Universal Robots PolyScope program: AdientTorsF_Eol21.urp

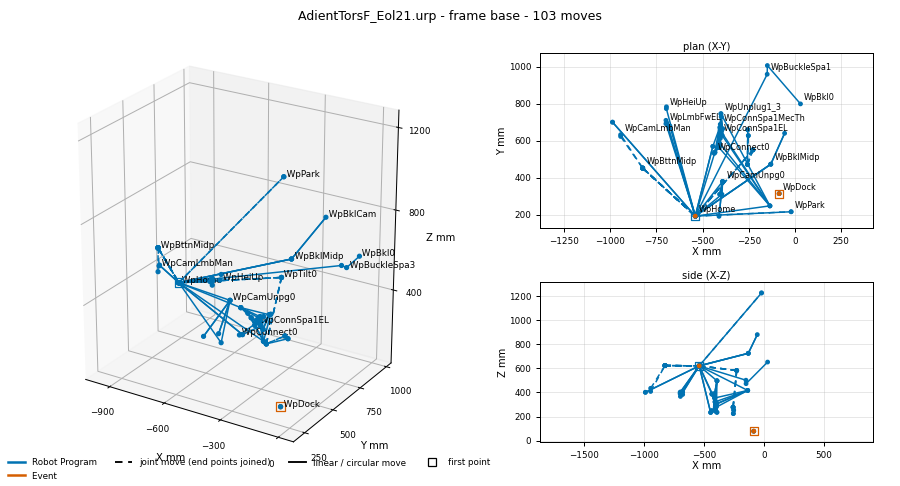
[picture p0: tool path of AdientTorsF_Eol21.urp in frame base, 103 of 155 moves have a stored position in this frame; points joined in program order, loops and branches not executed]
Program AdientTorsF_Eol21 (installation=EOL_21 directory=/programs createdIn=3.5.1 lastSavedIn=5.26.0 robotSerialNumber=20265101890)
Calibrated DH parameters: a=[0.000035, -0.496948, -0.566193, -0.00002, -0.00001, 0]; d=[0.180707, 184.637728, -195.556152, 11.09222, 0.119882, 0.115586]; alpha=[1.570552, -0.001939, 0.006964, 1.570414, -1.570475, 0]; deltaTheta=[0, -0.624231, 6.773924, 0.133492, -0.000002, 0]
InitVariablesNode variables(variable(name=Abort, expression=False), variable(name=AdapterReady, expression=False), variable(name=CMD_Heartbt_i1, expression=0), variable(name=CMD_Program_i1, expression=0), variable(name=CMD_Reserve_i1, expression=0), variable(name=CMD_Timeout_i1, expression=0), variable(name=CamCorrectnOK, expression=0), variable(name=DEBUG, expression=False), variable(name=D_rel, expression=p[0,0,0,0,0,0]), variable(name=EvtBeep, expression=False), variable(name=EvtDock, expression=0), variable(name=Mute, expression=False), variable(name=P_ini, expression=get_actual_tcp_pose()), variable(name=Parking, expression=0), variable(name=ProgExe, expression=0), variable(name=PusherPosFt, expression=0), variable(name=PusherReturn, expression=True), variable(name=STS_Heartbeat, expression=False), variable(name=STS_Progress, expression=0), variable(name=STS_Reservation, expression=0), variable(name=SetCameraProg, expression=0), variable(name=T_KeepReservtn, expression=0), variable(name=Tilt_PV, expression=0))
BeforeStart
  SuppressedNode
    DEBUG := True
  'SW version, to be used to track changes and keep sync of all stations'
  SW_Ver := 1.0
  Folder Scripts [hidden by the author, left out]
  Folder Avoid guidance screen
    Wp := get_actual_tcp_pose()
    MoveJ speed 120 deg/s, acceleration 500 deg/s^2 (useActiveTCP=true optimoveEnabled=false optiMoveSpeed=0.3 optiMoveAcceleration=0.09) feature=Base
      Waypoint Variable (Variable): variable=Wp
  Call GripperOpen
  GoToHome := True
  Script: socket_open("127.0.0.1",30001)
Robot Program (runOnlyOnce=false)
  Folder Execute Program
    Folder Init
      Wait Condition expression=EvtDock≤0
      Folder Verify Adapter ready
        If Di_Docked or AI_Gripper<(ivGripSensOpen+0.3)
          AdapterReady := False
      Folder Go to home pos automatically
        If GoToHome and  not AdapterReady
          Wait Sleep waitTime=1
          If InRange(P_Flange[0],-1,-0.2) and InRange(P_Flange[1],-0.5,0.5) and InRange(P_Flange[2],0.3,1)
            If AdapterDocked or DEBUG or (AI_Gripper<(ivGripSensOpen+0.3))
              MoveJ speed 120 deg/s, acceleration 500 deg/s^2 (useActiveTCP=false positionType=JointAngles optimoveEnabled=false optiMoveSpeed=0.3 optiMoveAcceleration=0.09) tcp=t0_Flange; feature=Base
                Waypoint WpHome: TCP in base x=-539.74 y=192.879 z=621.496 mm, rx=3.1416 ry=0 rz=0 rad; joints [177.915, -76.399, -107.627, -86.021, 90.391, 88.106] deg
            Else 
              Popup Error (haltProgram=false message=Adapter must be docked inputType=Text)
              Halt
          ElseIf AtParkPos
            MoveJ speed 120 deg/s, acceleration 500 deg/s^2 (useActiveTCP=false positionType=JointAngles optimoveEnabled=false optiMoveSpeed=0.3 optiMoveAcceleration=0.09) tcp=t0_Flange; feature=Base
              Waypoint WpPark: TCP in base x=-21.021 y=216.43 z=1228.484 mm, rx=-2.2794 ry=-2.1557 rz=0.0038 rad; joints [148.842, -80.043, -21.696, -168.004, 90.169, -28.26] deg
          Else 
            Popup Error (haltProgram=false message=Illegal position. Adjust arm to open space in front of the backrest, or [Move]->[Home] inputType=Text)
            Halt
        GoToHome := False
      If DEBUG
        'Popup window with program selection'
        ProgExe :=  (valueSource=Operator message=Program number? valueType=Integer)
      If ProgExe>0
        Folder Init
          Mute := False
          Wait Condition expression=not GoToHome
          If not In(ProgExe,[11,12,13,14])
            AdapterReady := False
    Folder Programs
      If InRange(ProgExe,1,99)
        Folder Undock
          If In(ProgExe,[11])
            Script: Report(1)
            If not AdapterReady
              Folder AtHome? [hidden by the author, left out]
              If Progress_run() and  not AdapterDocked
                Script: Report(94)
              If Progress_run()
                Folder Undock
                  MoveL speed 1000 mm/s, acceleration 3000 mm/s^2 (useActiveTCP=false optimoveEnabled=false optiMoveSpeed=0.3 optiMoveAcceleration=0.09) tcp=t2_Gripper; feature=Base
                    Call GripperOpenQuick
                    Wp := pose_trans(WpDock, p[0,0.175,-0.1,0,0,0])
                    Waypoint Variable (Variable): motionParameters(blendRadius=0.05); variable=Wp
                    Call GripperOpen
                    Wp := pose_trans(WpDock, p[0,0.075,0.01,0,0,0])
                    Waypoint Variable (Variable): motionParameters(blendRadius=0.01); variable=Wp
                    Wp := pose_trans(WpDock, p[0,0.055,0,0,0,0])
                    Waypoint Variable (Variable): motionParameters(blendRadius=0.01); variable=Wp
                    Waypoint WpDock: TCP in base x=-85.659 y=314.493 z=77.7 mm, rx=1.8875 ry=-1.8567 rz=-0.5938 rad; joints [149.519, -78.77, -155.163, -4.834, 107.001, 153.83] deg
                    Call GripperClose
                    Wp := pose_trans(WpDock, p[0,0.25,0,0,0,0])
                    Waypoint Variable (Variable): variable=Wp
                  AdapterReady := True
                  Script: Report(50)
            Else 
              Script: Report(50)
        Folder Connect
          If In(ProgExe,[12,13,14])
            Script: Report(1)
            PusherPosDev := 0
            MeasHeight := 0
            If not AdapterReady
              Folder AtHome? [hidden by the author, left out]
              If Progress_run() and  not AdapterDocked
                Script: Report(94)
            If Progress_run()
              Folder Length measure with pusher (mechanical seat)
                If In(ProgExe,[13])
                  Set DigitalOutput pin=Do_PusherReturn; digitalValue=0
                  Set DigitalOutput pin=Do_PusherWork; digitalValue=1
                Else 
                  PusherReturn := True
              Folder Undock
                If not AdapterReady
                  MoveL speed 1000 mm/s, acceleration 3000 mm/s^2 (useActiveTCP=false optimoveEnabled=false optiMoveSpeed=0.3 optiMoveAcceleration=0.09) tcp=t2_Gripper; feature=Base
                    Call GripperOpenQuick
                    Wp := pose_trans(WpDock, p[0,0.175,-0.1,0,0,0])
                    Waypoint Variable (Variable): motionParameters(blendRadius=0.05); variable=Wp
                    Call GripperOpen
                    Wp := pose_trans(WpDock, p[0,0.075,0.01,0,0,0])
                    Waypoint Variable (Variable): motionParameters(blendRadius=0.01); variable=Wp
                    Wp := pose_trans(WpDock, p[0,0.055,0,0,0,0])
                    Waypoint Variable (Variable): motionParameters(blendRadius=0.01); variable=Wp
                    Waypoint WpDock: TCP in base x=-85.659 y=314.493 z=77.7 mm, rx=1.8875 ry=-1.8567 rz=-0.5938 rad; joints [149.519, -78.77, -155.163, -4.834, 107.001, 153.83] deg
                    Call GripperClose
                    Wp := pose_trans(WpDock, p[0,0.25,0,0,0,0])
                    Waypoint Variable (Variable): variable=Wp
                AdapterReady := False
                Script: Report(2)
              CamCorrection := p[0,0,0,0,0,0]
              SuppressedNode
                Folder Camera
                  MoveL speed 1000 mm/s, acceleration 3000 mm/s^2 (useActiveTCP=false optimoveEnabled=false optiMoveSpeed=0.3 optiMoveAcceleration=0.09) tcp=t0_Flange; feature=Base
                    If In(ProgExe,[12,13])
                      SetCameraProg := 12
                      Waypoint WpCamCon0: motionParameters(blendRadius=0.05); TCP in base x=-326.648 y=291.698 z=338.41 mm, rx=2.1948 ry=2.1949 rz=-0.0575 rad; joints [160.702, -71.24, -141.099, -58.684, 93.132, -18.987] deg
                      Waypoint WpCamConSpa1: TCP in base x=-326.648 y=416.698 z=338.41 mm, rx=2.1948 ry=2.1949 rz=-0.0575 rad; joints [146.583, -82.407, -133.037, -56.241, 92.784, -33.102] deg
                    If In(ProgExe,[14])
                      SetCameraProg := ProgExe
                      Waypoint WpCamCon0: motionParameters(blendRadius=0.05); TCP in base x=-326.648 y=291.698 z=338.41 mm, rx=2.1948 ry=2.1949 rz=-0.0575 rad; joints [160.702, -71.24, -141.099, -58.684, 93.132, -18.987] deg
                      Waypoint WpCamConSpa3: TCP in base x=-370.516 y=382.662 z=354.732 mm, rx=-2.2214 ry=-2.2215 rz=0 rad; joints [153.025, -81.286, -132.366, -56.394, 90.281, -26.621] deg
                  Call CamAcquire
                  CamCorrection := p[CamData[0],CamData[1]*-0.5,CamData[1],0,0,0]
            CamCorrectnOK := ProgExe
            If In(ProgExe,[13])
              Timer (action=Reset) variable=T_Timeout
              Timer (action=Start) variable=T_Timeout
              Wait Condition expression=(PusherPosStable and InRange(PusherPos-ivPusherSeatRef,-15,15)) or T_Timeout>10
              PusherPosDev := PusherPos-ivPusherSeatRef
              If PusherPosStable and InRange(PusherPosDev,-15,15)
                'continue'
              Else 
                CamCorrectnOK := 0
                'CamCorrectionOK is also used as pusher measurement result'
            If Progress_run() and CamCorrectnOK≠ProgExe
              EvtDock := 1
              Wait Condition expression=EvtDock≤0
              Script: Report(91)
            If Progress_run() and ProgExe≟13
              'Wait handle catch done'
              Script: Report(3)
              Timer (action=Reset) variable=T_Timeout
              Timer (action=Start) variable=T_Timeout
              Wait Condition expression=Flags[12] or T_Timeout>10 or DEBUG
              If Flags[12] or DEBUG
                'ok'
              Else 
                Script: Report(98)
            If Progress_run() and  not Di_LiftDown
              EvtDock := 1
              Wait Condition expression=EvtDock≤0
              AdapterReady := False
              Script: Report(92)
            Folder Connect
              If Progress_run()
                Script: Report(4)
                Set NoAction tcp=t2_Gripper
                MoveL speed 1000 mm/s, acceleration 3000 mm/s^2 (useActiveTCP=false optimoveEnabled=false optiMoveSpeed=0.3 optiMoveAcceleration=0.09) tcp=t2_Gripper; feature=Base
                  Waypoint WpConnect0: TCP in base x=-437.091 y=531.932 z=249.935 mm, rx=3.1416 ry=0 rz=0 rad; joints [167.745, -81.605, -135.899, -52.542, 90.261, 78.118] deg; TCP offset x=0 y=-260 z=74 mm, rx=0 ry=0 rz=0 rad
                  If False
                    '30mm below connector, guides aligned (Y +-10mm)'
                    Waypoint WpConnSpa1EL: TCP in base x=-406.193 y=631.366 z=278.599 mm, rx=3.1251 ry=-0.0345 rz=0.0169 rad; joints [155.804, -83.836, -129.752, -57.368, 90.869, 67.396] deg; TCP offset x=0 y=-260 z=74 mm, rx=0 ry=0 rz=0 rad
                    Waypoint WpConnSpa1Mec: TCP in base x=-404.448 y=625.534 z=295.592 mm, rx=3.0512 ry=-0.0001 rz=0 rad; joints [154.483, -81.409, -127.32, -63.499, 94.969, 64.697] deg; TCP offset x=0 y=-260 z=74 mm, rx=0 ry=0 rz=0 rad
                    Waypoint WpConnSpa3: TCP in base x=-397.516 y=650.604 z=285.207 mm, rx=3.1416 ry=0 rz=0 rad; joints [153.476, -83.698, -129.812, -56.508, 90.26, 63.812] deg; TCP offset x=0 y=-260 z=74 mm, rx=0 ry=0 rz=0 rad
                    'Touching the plug from below, seat is in assy(3 pumps from topmost)'
                    Waypoint WpConnSpa1MecTh: TCP in base x=-404.456 y=689.742 z=287.147 mm, rx=3.0512 ry=-0.0001 rz=0 rad; joints [148.645, -86.649, -123.608, -62.436, 94.705, 58.848] deg; TCP offset x=0 y=-260 z=74 mm, rx=0 ry=0 rz=0 rad
                  If In(ProgExe,[12])
                    Wp := WpConnSpa1EL
                  If In(ProgExe,[13])
                    'adjust angle mechanical'
                    Wp0 := pose_add(WpConnSpa1MecTh,p[0,PusherPosDev/1000,-0.025,0,0,0])
                    Waypoint Variable (Variable): variable=Wp0
                    Force Frame feature=Joint_6_name; selection=[0, 0, 1, 0, 0, 0]; wrench=[0, 0, -30, -0.5, 0, 0]; limitsForce=[0.15, 0.15, 0.1, 0.087266, 1.047198, 1.047198]; limitsMotion=[0.1, 0.1, 0.1, 0.349066, 0.349066, 0.349066]
                      Wait Sleep waitTime=0.5
                    Force Frame feature=Joint_6_name; selection=[0, 0, 1, 0, 0, 0]; wrench=[0, 0, -10, -0.5, 0, 0]; limitsForce=[0.15, 0.15, 0.002, 0.087266, 1.047198, 1.047198]; limitsMotion=[0.1, 0.1, 0.1, 0.349066, 0.349066, 0.349066]
                      Wait Sleep waitTime=0.5
                    Wp := get_actual_tcp_pose()
                    MeasHeight := (Wp[2]-WpConnSpa1MecTh[2])*1000
                    MoveDirectionNode expression=[0.0,1.0,0.2]; feature=Joint_6_name
                      Until DISTANCE (allowActions=false deceleration=3 distanceNodeType=STOP) Distance=0.07; motionParameters(blendRadius=0)
                    Wp := pose_add(WpConnSpa1Mec,p[0,PusherPosDev/1000,0,0,0,0])
                    CorrMechSeat := p[0,0,0,0,0,0]
                    If MeasHeight>0
                      Script: CorrMechSeat[1]=Calibrate(MeasHeight,0,17,0,-7)/1000
                      Script: CorrMechSeat[2]=Calibrate(MeasHeight,0,17,0,26)/1000
                      Script: CorrMechSeat[3]=Calibrate(MeasHeight,0,17,0,-0.129)
                    Else 
                      Script: CorrMechSeat[1]=Calibrate(MeasHeight,-13,0,7,0)/1000
                      Script: CorrMechSeat[2]=Calibrate(MeasHeight,-13,0,-19,0)/1000
                      Script: CorrMechSeat[3]=Calibrate(MeasHeight,-13,0,0.053,0)
                    Wp := pose_add(Wp,CorrMechSeat)
                  If In(ProgExe,[14])
                    Wp := WpConnSpa3
                  Waypoint Variable (Variable): variable=Wp
                Force Frame feature=Joint_6_name; selection=[0, 0, 1, 0, 0, 0]; wrench=[0, 0, -30, 0, 0, 0]; limitsForce=[0.15, 0.15, 0.1, 1.047198, 1.047198, 1.047198]; limitsMotion=[0.1, 0.1, 0.1, 0.349066, 0.349066, 0.349066]
                  Wait Sleep waitTime=1
                Force Frame feature=Joint_6_name; selection=[1, 0, 1, 0, 0, 0]; wrench=[0, 0, -30, 0, 0, 0]; limitsForce=[0.15, 0.15, 0.05, 1.047198, 1.047198, 1.047198]; limitsMotion=[0.1, 0.1, 0.1, 0.349066, 0.349066, 0.349066]
                  Wait Sleep waitTime=0.5
                'position ok, not checked for mechanical seat'
                If InRange(Wp[2]+0.03-P_act[2],-0.015,0.015) or ProgExe≟13
                  'ok'
                Else 
                  EvtDock := 2
                  Wait Condition expression=EvtDock≤0
                  Script: Report(96)
              If Progress_run()
                Force Frame feature=Joint_6_name; selection=[0, 1, 0, 0, 0, 0]; wrench=[0, -60, -10, 0, 0, 0]; limitsForce=[0.15, 0.05, 0.01, 1.047198, 1.047198, 1.047198]; limitsMotion=[0.1, 0.1, 0.1, 0.349066, 0.349066, 0.349066]
                  Wait Sleep waitTime=1
                MoveL speed 1000 mm/s, acceleration 3000 mm/s^2 (useActiveTCP=true optimoveEnabled=false optiMoveSpeed=0.3 optiMoveAcceleration=0.09) feature=Base
                  Wp := pose_trans(P_act, p[0,0.005,0,0,0,0])
                  Waypoint Variable (Variable): variable=Wp
                Call GripperOpen
                Force Frame feature=Joint_6_name; selection=[0, 1, 0, 0, 0, 0]; wrench=[0, -60, -10, 0, 0, 0]; limitsForce=[0.15, 0.1, 0.01, 1.047198, 1.047198, 1.047198]; limitsMotion=[0.1, 0.1, 0.1, 0.349066, 0.349066, 0.349066]
                  Wait Sleep waitTime=1
                  Script: Report(5)
                  MoveL speed 500 mm/s, acceleration 2000 mm/s^2 (useActiveTCP=true optimoveEnabled=false optiMoveSpeed=0.3 optiMoveAcceleration=0.09) feature=Base
                    Wp0 := get_actual_tcp_pose()
                    Wp := pose_trans(Wp0, p[0,0,0,0,0,0.07])
                    Waypoint Variable (Variable): variable=Wp
                    Wp := pose_trans(Wp0, p[0,0,0,0,0,-0.07])
                    Waypoint Variable (Variable): variable=Wp
                    Waypoint Variable (Variable): variable=Wp0
                    Wp := pose_trans(Wp0, p[0,0,0.01,0,0,0])
                    Waypoint Variable (Variable): variable=Wp
                    Waypoint Variable (Variable): variable=Wp0
                MoveL speed 1000 mm/s, acceleration 3000 mm/s^2 (useActiveTCP=true optimoveEnabled=false optiMoveSpeed=0.3 optiMoveAcceleration=0.09) feature=Base
                  Wp0 := get_actual_tcp_pose()
                  Wp := pose_trans(Wp0, p[0,0.015,0,0,0,0])
                  Waypoint Variable (Variable): variable=Wp
                Force Frame feature=Joint_6_name; selection=[0, 1, 0, 0, 0, 0]; wrench=[0, -60, 0, 0, 0, 0]; limitsForce=[0.15, 0.5, 0.15, 1.047198, 1.047198, 1.047198]; limitsMotion=[0.1, 0.1, 0.1, 0.349066, 0.349066, 0.349066]
                  Wait Sleep waitTime=0.5
                Script: Report(6)
                Timer (action=Reset) variable=T_Timeout
                Timer (action=Start) variable=T_Timeout
                Folder Test switch pin, retreat on fail
                  Wait Condition expression=Flags[0] or T_Timeout>10 or DEBUG
                  If not Flags[0] and  not DEBUG
                    EvtDock := 2
                    Wait Condition expression=EvtDock≤0
                    Script: Report(95)
            If Progress_run()
              MoveL speed 1000 mm/s, acceleration 3000 mm/s^2 (useActiveTCP=false optimoveEnabled=false optiMoveSpeed=0.3 optiMoveAcceleration=0.09) tcp=t0_Flange; feature=Base
                Set NoAction tcp=t0_Flange
                P_act := get_actual_tcp_pose()
                Wp := pose_trans(P_act, p[0,0.1,0,0,0,0])
                Waypoint Variable (Variable): motionParameters(blendRadius=0.05); variable=Wp
                Wp := pose_trans(Wp, p[-0.15,0.1,-0.2,0,0.5,0])
                Waypoint Variable (Variable): motionParameters(blendRadius=0.05); variable=Wp
                Waypoint WpHome: TCP in base x=-539.74 y=192.879 z=621.496 mm, rx=3.1416 ry=0 rz=0 rad; joints [177.915, -76.399, -107.627, -86.021, 90.391, 88.106] deg
              Script: Report(50)
        Folder Buckle
          If In(ProgExe,[15,16])
            Script: Report(1)
            Folder AtHome? [hidden by the author, left out]
            If Progress_run()
              Call GripperCloseQuick
              Folder Camera
                SetCameraProg := ProgExe
                MoveL speed 1000 mm/s, acceleration 3000 mm/s^2 (useActiveTCP=false optimoveEnabled=false optiMoveSpeed=0.3 optiMoveAcceleration=0.09) tcp=t0_Flange; feature=Base
                  Waypoint WpBklMidp: motionParameters(blendRadius=0.05); TCP in base x=-131.026 y=473.792 z=726.036 mm, rx=-2.1821 ry=2.2601 rz=0 rad; joints [126.005, -68.539, -102.415, -99.065, 90.386, 128.091] deg
                  Waypoint WpBklCam: TCP in base x=-56.214 y=641.103 z=881.577 mm, rx=-1.8636 ry=0.3608 rz=-1.6302 rad; joints [121.325, -95.448, -62.678, -192.662, 15.525, 118.92] deg
                Call GripperClose
                Call CamAcquire
                Call CamCalculateCorectnPlane
                If CamCorrectnOK≟ProgExe and InRange(CamCorrection[1],-0.05,0.05) and InRange(CamCorrection[2],-0.03,0.03)
                  'empty'
                Else 
                  CamCorrectnOK := 0
                  MoveL speed 1000 mm/s, acceleration 3000 mm/s^2 (useActiveTCP=false optimoveEnabled=false optiMoveSpeed=0.3 optiMoveAcceleration=0.09) tcp=t0_Flange; feature=Base
                    Waypoint WpBklMidp: motionParameters(blendRadius=0.05); TCP in base x=-131.026 y=473.792 z=726.036 mm, rx=-2.1821 ry=2.2601 rz=0 rad; joints [126.005, -68.539, -102.415, -99.065, 90.386, 128.091] deg
                    Waypoint WpHome: TCP in base x=-539.74 y=192.879 z=621.496 mm, rx=3.1416 ry=0 rz=0 rad; joints [177.915, -76.399, -107.627, -86.021, 90.391, 88.106] deg
                  Script: Report(91)
              If CamCorrectnOK≟ProgExe
                Folder Insert
                  MoveL speed 1000 mm/s, acceleration 3000 mm/s^2 (useActiveTCP=false optimoveEnabled=false optiMoveSpeed=0.3 optiMoveAcceleration=0.09) tcp=t3_Blade; feature=Base
                    If False
                      'must be set with blade ca one half into buckle slot'
                      Waypoint WpBuckleSpa1: TCP in base x=-150.458 y=960.619 z=502.148 mm, rx=-2.7056 ry=-0.0003 rz=0.0018 rad; joints [103.392, -102.167, -91.983, -51.502, 84.645, 12.49] deg; TCP offset x=-134 y=-56 z=118 mm, rx=0 ry=0 rz=0 rad
                      Waypoint WpBuckleSpa3: TCP in base x=-149.61 y=1007.832 z=473.301 mm, rx=-2.5307 ry=0 rz=0 rad; joints [103.075, -106.712, -94.104, -34.951, 82.628, 11.124] deg
                    If ProgExe≟15
                      Wp := WpBuckleSpa1
                    If ProgExe≟16
                      Wp := WpBuckleSpa3
                    Wp0 := pose_trans(Wp,p[0,0,-0.02,0,0,0])
                    Wp0 := pose_add(Wp0,Base_w_correctn)
                    Waypoint WpBkl0: motionParameters(blendRadius=0.05); TCP in base x=29.678 y=800.175 z=653.181 mm, rx=-2.8405 ry=-0.1319 rz=-1.2182 rad; joints [106.833, -94.053, -71.668, -115.292, 44.916, 16.097] deg
                    Waypoint Variable (Variable): variable=Wp0
                  Script: Report(5)
                  Timer (action=Reset) variable=T_Timeout
                  Timer (action=Start) variable=T_Timeout
                  Wait Condition expression=Flags[8] or Abort or DEBUG  or T_Timeout>25
                  If Flags[8] or DEBUG
                    Script: Report(6)
                    Set NoAction tcp=t3_Blade
                    Force Frame feature=Joint_6_name; selection=[0, 0, 1, 0, 0, 0]; wrench=[0, 0, 15, 0, 0, 0]; limitsForce=[0.15, 0.15, 0.15, 1.047198, 1.047198, 1.047198]; limitsMotion=[0.1, 0.1, 0.1, 0.349066, 0.349066, 0.349066]
                      Wait Sleep waitTime=1
                    If not Flags[9] and  not Abort
                      MoveL speed 50 mm/s, acceleration 500 mm/s^2 (useActiveTCP=false optimoveEnabled=false optiMoveSpeed=0.3 optiMoveAcceleration=0.09) tcp=t3_Blade; feature=Base
                        Waypoint Variable (Variable): variable=Wp
                      Force Frame feature=Joint_6_name; selection=[1, 1, 1, 0, 0, 0]; wrench=[0, 0, 50, 0, 0, 0]; limitsForce=[0.15, 0.15, 0.25, 1.047198, 1.047198, 1.047198]; limitsMotion=[0.1, 0.1, 0.1, 0.349066, 0.349066, 0.349066]
                        Wait Sleep waitTime=1.5
                    If not Flags[9] and  not Abort
                      MoveL speed 50 mm/s, acceleration 500 mm/s^2 (useActiveTCP=false optimoveEnabled=false optiMoveSpeed=0.3 optiMoveAcceleration=0.09) tcp=t3_Blade; feature=Base
                        Waypoint Variable (Variable): variable=Wp
                      Force Frame feature=Joint_6_name; selection=[1, 1, 1, 0, 0, 0]; wrench=[0, 0, 50, 0, 0, 0]; limitsForce=[0.15, 0.15, 0.25, 1.047198, 1.047198, 1.047198]; limitsMotion=[0.1, 0.1, 0.1, 0.349066, 0.349066, 0.349066]
                        Wait Sleep waitTime=1.5
                    If not Flags[9] and  not Abort
                      MoveL speed 50 mm/s, acceleration 500 mm/s^2 (useActiveTCP=false optimoveEnabled=false optiMoveSpeed=0.3 optiMoveAcceleration=0.09) tcp=t3_Blade; feature=Base
                        Waypoint Variable (Variable): variable=Wp
                      Force Frame feature=Joint_6_name; selection=[1, 1, 1, 0, 0, 0]; wrench=[0, 0, 50, 0, 0, 0]; limitsForce=[0.15, 0.15, 0.25, 1.047198, 1.047198, 1.047198]; limitsMotion=[0.1, 0.1, 0.1, 0.349066, 0.349066, 0.349066]
                        Wait Sleep waitTime=1.5
                  MoveL speed 1000 mm/s, acceleration 3000 mm/s^2 (useActiveTCP=false optimoveEnabled=false optiMoveSpeed=0.3 optiMoveAcceleration=0.09) tcp=t3_Blade; feature=Base
                    Waypoint Variable (Variable): variable=Wp
                    MoveDirectionNode (selectedDirection=ZMinus) feature=Joint_6_name
                      Until DISTANCE (allowActions=false deceleration=3 distanceNodeType=STOP) Distance=0.02; motionParameters(blendRadius=0)
                  MoveL speed 1000 mm/s, acceleration 3000 mm/s^2 (useActiveTCP=false optimoveEnabled=false optiMoveSpeed=0.3 optiMoveAcceleration=0.09) tcp=t0_Flange; feature=Base
                    Waypoint WpBklMidp: motionParameters(blendRadius=0.05); TCP in base x=-131.026 y=473.792 z=726.036 mm, rx=-2.1821 ry=2.2601 rz=0 rad; joints [126.005, -68.539, -102.415, -99.065, 90.386, 128.091] deg
                    Waypoint WpHome: TCP in base x=-539.74 y=192.879 z=621.496 mm, rx=3.1416 ry=0 rz=0 rad; joints [177.915, -76.399, -107.627, -86.021, 90.391, 88.106] deg
                  If Progress_check()≥6
                    Script: Report(50)
                  Else 
                    Script: Report(95)
        Folder Disconnect
          If In(ProgExe,[21,22,23])
            Script: Report(1)
            Folder AtHome? [hidden by the author, left out]
            If Progress_run()
              If In(ProgExe,[21])
                SetCameraProg := ProgExe
                MoveL speed 1000 mm/s, acceleration 3000 mm/s^2 (useActiveTCP=false optimoveEnabled=false optiMoveSpeed=0.3 optiMoveAcceleration=0.09) tcp=t0_Flange; feature=Base
                  Waypoint WpCamUnpg0: motionParameters(blendRadius=0.05); TCP in base x=-391.776 y=380.411 z=497.114 mm, rx=2.149 ry=-2.149 rz=0.1503 rad; joints [152.651, -76.876, -119.272, -77.538, 97.454, 152.641] deg
                  Waypoint WpCamUnplgSpa1: TCP in base x=-408.404 y=310.844 z=356.503 mm, rx=2.149 ry=-2.149 rz=0.1503 rad; joints [160.519, -79.837, -132.767, -60.055, 97.826, 160.666] deg
              If In(ProgExe,[22])
                SetCameraProg := ProgExe
                MoveL speed 1000 mm/s, acceleration 3000 mm/s^2 (useActiveTCP=false optimoveEnabled=false optiMoveSpeed=0.3 optiMoveAcceleration=0.09) tcp=t0_Flange; feature=Base
                  Waypoint WpCamUnpg0: motionParameters(blendRadius=0.05); TCP in base x=-391.776 y=380.411 z=497.114 mm, rx=2.149 ry=-2.149 rz=0.1503 rad; joints [152.651, -76.876, -119.272, -77.538, 97.454, 152.641] deg
                  Waypoint WpCamUnplgSpa1M: TCP in base x=-411.184 y=191.542 z=392.404 mm, rx=2.149 ry=-2.149 rz=0.1503 rad; joints [175.142, -70.201, -135.712, -64.745, 98.291, 175.397] deg
              If In(ProgExe,[23])
                SetCameraProg := ProgExe
                MoveL speed 1000 mm/s, acceleration 3000 mm/s^2 (useActiveTCP=false optimoveEnabled=false optiMoveSpeed=0.3 optiMoveAcceleration=0.09) tcp=t0_Flange; feature=Base
                  Waypoint WpCamUnpg0: motionParameters(blendRadius=0.05); TCP in base x=-391.776 y=380.411 z=497.114 mm, rx=2.149 ry=-2.149 rz=0.1503 rad; joints [152.651, -76.876, -119.272, -77.538, 97.454, 152.641] deg
                  Waypoint WpCamUnpgSpa3: TCP in base x=-395.254 y=310.844 z=314.879 mm, rx=2.2011 ry=-2.2011 rz=0.0444 rad; joints [161.28, -81.245, -137.148, -52.352, 92.432, 161.627] deg; TCP offset x=0 y=0 z=0 mm, rx=0 ry=0 rz=0 rad
              Call CamAcquire
              Call CamCalculateCorectnPlane
            If Progress_run() and CamCorrectnOK≠ProgExe
              MoveL speed 1000 mm/s, acceleration 3000 mm/s^2 (useActiveTCP=false optimoveEnabled=false optiMoveSpeed=0.3 optiMoveAcceleration=0.09) tcp=t0_Flange; feature=Base
                Waypoint WpHome: TCP in base x=-539.74 y=192.879 z=621.496 mm, rx=3.1416 ry=0 rz=0 rad; joints [177.915, -76.399, -107.627, -86.021, 90.391, 88.106] deg
              Script: Report(91)
            If Progress_run()
              Call GripperOpenQuick
              Folder Disconnect
                If In(ProgExe,[21])
                  MoveL speed 1000 mm/s, acceleration 3000 mm/s^2 (useActiveTCP=false optimoveEnabled=false optiMoveSpeed=0.3 optiMoveAcceleration=0.09) tcp=t2_Gripper; feature=Base_w_correctn
                    Waypoint WpUnplg_0: motionParameters(blendRadius=0.05); TCP in base x=-135.864 y=248.289 z=416.995 mm, rx=2.2887 ry=-2.152 rz=0.0002 rad; joints [171.613, -65.804, -127.743, -76.476, 90.37, 168.318] deg; TCP offset x=0 y=-260 z=74 mm, rx=0 ry=0 rz=0 rad
                    Call GripperOpen
                    Waypoint WpUnplug1_1: motionParameters(blendRadius=0.05); TCP in base x=-407.93 y=586.737 z=321.99 mm, rx=2.6768 ry=0 rz=0 rad; joints [149.589, -81.15, -114.014, -89.039, 113.125, 56.858] deg
                    Waypoint WpUnplug1_2: motionParameters(blendRadius=0.05); TCP in base x=-403.747 y=662.579 z=254.257 mm, rx=2.6768 ry=0 rz=0 rad; joints [143.353, -88.891, -113.69, -84.034, 111.445, 50.41] deg
                    Waypoint WpUnplug1_3: TCP in base x=-400.842 y=747.152 z=275.935 mm, rx=3.131 ry=-0.0006 rz=0.0001 rad; joints [145.117, -91.643, -122.979, -55.744, 90.742, 55.469] deg
                If In(ProgExe,[22])
                  MoveL speed 1000 mm/s, acceleration 3000 mm/s^2 (useActiveTCP=false optimoveEnabled=false optiMoveSpeed=0.3 optiMoveAcceleration=0.09) tcp=t2_Gripper; feature=Base_w_correctn
                    Waypoint WpUnplg_0: motionParameters(blendRadius=0.05); TCP in base x=-135.864 y=248.289 z=416.995 mm, rx=2.2887 ry=-2.152 rz=0.0002 rad; joints [171.613, -65.804, -127.743, -76.476, 90.37, 168.318] deg
                    Call GripperOpen
                    Waypoint WpUnplug_1_1M: motionParameters(blendRadius=0.04); TCP in base x=-411.15 y=563.75 z=353.982 mm, rx=2.6768 ry=0 rz=0 rad; joints [151.779, -78.91, -112.719, -91.677, 113.652, 59.149] deg
                    Waypoint WpUnplug1_2M: motionParameters(blendRadius=0.05); TCP in base x=-405.13 y=613.357 z=273.879 mm, rx=2.6768 ry=0 rz=0 rad; joints [147.213, -84.488, -116.009, -84.645, 112.511, 54.402] deg
                    Waypoint WpUnplg1_3M: TCP in base x=-404.987 y=658.915 z=299.047 mm, rx=3.0284 ry=-0.0005 rz=0.0001 rad; joints [150.936, -83.747, -124.113, -65.294, 95.966, 61.089] deg
                If In(ProgExe,[23])
                  MoveL speed 1000 mm/s, acceleration 3000 mm/s^2 (useActiveTCP=false optimoveEnabled=false optiMoveSpeed=0.3 optiMoveAcceleration=0.09) tcp=t2_Gripper; feature=Base_w_correctn
                    Waypoint WpUnplg_0: motionParameters(blendRadius=0.05); TCP in base x=-135.864 y=248.289 z=416.995 mm, rx=2.2887 ry=-2.152 rz=0.0002 rad; joints [171.613, -65.804, -127.743, -76.476, 90.37, 168.318] deg
                    Call GripperOpen
                    Waypoint WpUnplg3_2: motionParameters(blendRadius=0.05); TCP in base x=-395.147 y=630.549 z=306.611 mm, rx=2.7856 ry=0 rz=0 rad; joints [147.756, -82.381, -117.1, -81.702, 107.51, 56.252] deg
                    Waypoint WpUnplg3_3: motionParameters(blendRadius=0.025); TCP in base x=-392.142 y=665.322 z=234.916 mm, rx=2.7856 ry=0 rz=0 rad; joints [144.771, -87.891, -119.779, -74.386, 106.881, 53.244] deg
                    Waypoint WpUnplg3_4: TCP in base x=-399.107 y=730.4 z=281.046 mm, rx=3.1224 ry=0 rz=0 rad; joints [146.206, -89.918, -123.786, -56.919, 91.165, 56.529] deg
                Script: Report(20)
                Wait Condition expression=Flags[7] or DEBUG
              EvtDock := 2
              Wait Condition expression=EvtDock≤0
              If EvtDock<0
                If In(ProgExe,[21])
                  MoveL speed 1000 mm/s, acceleration 3000 mm/s^2 (useActiveTCP=false optimoveEnabled=false optiMoveSpeed=0.3 optiMoveAcceleration=0.09) tcp=t2_Gripper; feature=Base_w_correctn
                    Waypoint WpUnplug1_3: TCP in base x=-400.842 y=747.152 z=275.935 mm, rx=3.131 ry=-0.0006 rz=0.0001 rad; joints [145.117, -91.643, -122.979, -55.744, 90.742, 55.469] deg
                    Waypoint WpUnplug1_2: TCP in base x=-403.747 y=662.579 z=254.257 mm, rx=2.6768 ry=0 rz=0 rad; joints [143.353, -88.891, -113.69, -84.034, 111.445, 50.41] deg
                    Waypoint WpUnplug1_1: TCP in base x=-407.93 y=586.737 z=321.99 mm, rx=2.6768 ry=0 rz=0 rad; joints [149.589, -81.15, -114.014, -89.039, 113.125, 56.858] deg
                    Waypoint WpUnplug_1: TCP in base x=-433.594 y=537.985 z=386.664 mm, rx=3.1416 ry=0 rz=0 rad; joints [166.968, -73.547, -126.184, -70.315, 90.348, 77.251] deg
                If In(ProgExe,[22])
                  MoveL speed 1000 mm/s, acceleration 3000 mm/s^2 (useActiveTCP=false optimoveEnabled=false optiMoveSpeed=0.3 optiMoveAcceleration=0.09) tcp=t2_Gripper; feature=Base_w_correctn
                    Waypoint WpUnplg1_3M: TCP in base x=-404.987 y=658.915 z=299.047 mm, rx=3.0284 ry=-0.0005 rz=0.0001 rad; joints [150.936, -83.747, -124.113, -65.294, 95.966, 61.089] deg
                    Waypoint WpUnplug1_2M: TCP in base x=-405.13 y=613.357 z=273.879 mm, rx=2.6768 ry=0 rz=0 rad; joints [147.213, -84.488, -116.009, -84.645, 112.511, 54.402] deg
                    Waypoint WpUnplug_1_1M: TCP in base x=-411.15 y=563.75 z=353.982 mm, rx=2.6768 ry=0 rz=0 rad; joints [151.779, -78.91, -112.719, -91.677, 113.652, 59.149] deg
                    Waypoint WpUnplug_1: TCP in base x=-433.594 y=537.985 z=386.664 mm, rx=3.1416 ry=0 rz=0 rad; joints [166.968, -73.547, -126.184, -70.315, 90.348, 77.251] deg
                If In(ProgExe,[23])
                  MoveL speed 1000 mm/s, acceleration 3000 mm/s^2 (useActiveTCP=false optimoveEnabled=false optiMoveSpeed=0.3 optiMoveAcceleration=0.09) tcp=t2_Gripper; feature=Base_w_correctn
                    Waypoint WpUnplg3_4: TCP in base x=-399.107 y=730.4 z=281.046 mm, rx=3.1224 ry=0 rz=0 rad; joints [146.206, -89.918, -123.786, -56.919, 91.165, 56.529] deg
                    Waypoint WpUnplg3_3: TCP in base x=-392.142 y=665.322 z=234.916 mm, rx=2.7856 ry=0 rz=0 rad; joints [144.771, -87.891, -119.779, -74.386, 106.881, 53.244] deg
                    Waypoint WpUnplg3_2: motionParameters(blendRadius=0.05); TCP in base x=-395.147 y=630.549 z=306.611 mm, rx=2.7856 ry=0 rz=0 rad; joints [147.756, -82.381, -117.1, -81.702, 107.51, 56.252] deg
                    Waypoint WpUnplug_1: motionParameters(blendRadius=0.05); TCP in base x=-433.594 y=537.985 z=386.664 mm, rx=3.1416 ry=0 rz=0 rad; joints [166.968, -73.547, -126.184, -70.315, 90.348, 77.251] deg
                MoveL speed 1000 mm/s, acceleration 3000 mm/s^2 (useActiveTCP=false optimoveEnabled=false optiMoveSpeed=0.3 optiMoveAcceleration=0.09) tcp=t0_Flange; feature=Base
                  Waypoint WpHome: TCP in base x=-539.74 y=192.879 z=621.496 mm, rx=3.1416 ry=0 rz=0 rad; joints [177.915, -76.399, -107.627, -86.021, 90.391, 88.106] deg
                Script: Report(97)
            If Progress_run()
              Script: Report(50)
        Folder Buttons
          If In(ProgExe,[31,32,34])
            Script: Report(1)
            Call GripperCloseQuick
            Folder AtHome? [hidden by the author, left out]
            If Progress_run() and  not Di_SBR_X_Wp
              Script: Report(92)
            Folder Camera
              If Progress_run()
                If In(ProgExe,[31,32])
                  SetCameraProg := 32
                  MeasHeight := 0
                If In(ProgExe,[34])
                  SetCameraProg := 34
                MoveJ speed 120 deg/s, acceleration 500 deg/s^2 (useActiveTCP=false optimoveEnabled=false optiMoveSpeed=0.3 optiMoveAcceleration=0.09) tcp=t0_Flange; feature=Base
                  Waypoint WpBttnMidp: motionParameters(blendRadius=0.05); TCP in base x=-824.236 y=452.377 z=623.923 mm, rx=2.2214 ry=-2.2214 rz=0 rad; joints [161.838, -112.329, -68.535, -89.151, 90.318, 161.934] deg
                  Call GripperClose
                  If In(ProgExe,[34])
                    If False
                      Waypoint WpCamLmbMan: TCP in base x=-943.684 y=633.441 z=434.715 mm, rx=0.4666 ry=-3.0555 rz=0.0119 rad; joints [154.692, -134.904, -52.105, -80.844, 92.273, 227.473] deg
                    Wp := pose_add(WpCamLmbMan,p[0,0,MeasHeight/1000,0,0,0])
                    Waypoint Variable (Variable): variable=Wp
                  Else 
                    Waypoint WpCamLmbEL: TCP in base x=-943.684 y=623.984 z=408.727 mm, rx=0.4742 ry=-3.1055 rz=-0.0001 rad; joints [155.333, -135.057, -53.992, -80.965, 90.285, 228.08] deg
                Call CamAcquire
                Script: CamData[1]=CamData[1]-MeasHeight/1000
                Call CamCalculateCorectnPlane
            If Progress_run() and CamCorrectnOK≠ProgExe
              MoveJ speed 120 deg/s, acceleration 500 deg/s^2 (useActiveTCP=false positionType=JointAngles optimoveEnabled=false optiMoveSpeed=0.3 optiMoveAcceleration=0.09) tcp=t0_Flange; feature=Base
                Waypoint WpBttnMidp: motionParameters(blendRadius=0.05); TCP in base x=-824.236 y=452.377 z=623.923 mm, rx=2.2214 ry=-2.2214 rz=0 rad; joints [161.838, -112.329, -68.535, -89.151, 90.318, 161.934] deg
                Waypoint WpHome: TCP in base x=-539.74 y=192.879 z=621.496 mm, rx=3.1416 ry=0 rz=0 rad; joints [177.915, -76.399, -107.627, -86.021, 90.391, 88.106] deg
              Script: Report(91)
            Folder Lumbar
              If Progress_run()
                If In(ProgExe,[31,32])
                  Timer (action=Reset) variable=T_Timeout
                  Timer (action=Start) variable=T_Timeout
                  Script: Report(12)
                  Wait Condition expression=Flags[2] or T_Timeout>60 or DEBUG or Abort
                  If Flags[2] or DEBUG
                    MoveL speed 1000 mm/s, acceleration 3000 mm/s^2 (useActiveTCP=false optimoveEnabled=false optiMoveSpeed=0.3 optiMoveAcceleration=0.09) tcp=t4_Finger; feature=Base
                      Folder Press FW
                        If False
                          Waypoint WpLmbFwEL: TCP in base x=-698.714 y=692.998 z=390.507 mm, rx=0.3862 ry=-3.1106 rz=0.163 rad; joints [148.782, -134.738, -49.026, -89.82, 95.073, 224.534] deg; TCP offset x=-159 y=-58 z=70 mm, rx=0 ry=0 rz=0 rad
                        Wp := pose_trans(WpLmbFwEL, CamCorrection)
                        Waypoint Variable (Variable): variable=Wp
                        Force Frame feature=Joint_6_name; selection=[1, 0, 0, 0, 0, 0]; wrench=[-20, 10, -20, 0, 0, 0]; limitsForce=[0.05, 0.01, 0.05, 1.047198, 1.047198, 1.047198]; limitsMotion=[0.1, 0.1, 0.1, 0.349066, 0.349066, 0.349066]
                          Wait Sleep waitTime=0.7
                        ButtonPos := get_actual_tcp_pose()
                        Waypoint Variable (Variable): variable=Wp
                    Script: Report(3)
                  Else 
                    MoveJ speed 120 deg/s, acceleration 500 deg/s^2 (useActiveTCP=false optimoveEnabled=false optiMoveSpeed=0.3 optiMoveAcceleration=0.09) tcp=t0_Flange; feature=Base
                      Waypoint WpBttnMidp: motionParameters(blendRadius=0.05); TCP in base x=-824.236 y=452.377 z=623.923 mm, rx=2.2214 ry=-2.2214 rz=0 rad; joints [161.838, -112.329, -68.535, -89.151, 90.318, 161.934] deg
                      Waypoint WpHome: TCP in base x=-539.74 y=192.879 z=621.496 mm, rx=3.1416 ry=0 rz=0 rad; joints [177.915, -76.399, -107.627, -86.021, 90.391, 88.106] deg
                    Script: Report(95)
            Folder Multiring
              If Progress_run()
                If In(ProgExe,[32])
                  Timer (action=Reset) variable=T_Timeout
                  Timer (action=Start) variable=T_Timeout
                  Script: Report(11)
                  Wait Condition expression=Flags[1] or T_Timeout>60 or DEBUG or Abort
                  If Flags[1] or DEBUG
                    MoveL speed 1000 mm/s, acceleration 3000 mm/s^2 (useActiveTCP=false optimoveEnabled=false optiMoveSpeed=0.3 optiMoveAcceleration=0.09) tcp=t4_Finger; feature=Base
                      If False
                        Waypoint WpMultiringHi: TCP in base x=-677.239 y=680.361 z=403.46 mm, rx=0.3862 ry=-3.1106 rz=0.163 rad; joints [148.76, -131.638, -53.105, -88.842, 95.073, 224.524] deg; TCP offset x=-159 y=-58 z=70 mm, rx=0 ry=0 rz=0 rad
                        Waypoint WpMutiringLo: TCP in base x=-677.374 y=678.43 z=383.517 mm, rx=0.3862 ry=-3.1106 rz=0.163 rad; joints [148.847, -131.73, -54.956, -86.89, 95.076, 224.624] deg
                      Folder Press up
                        Wp0 := pose_add(WpMutiringLo,Base_w_correctn)
                        Wp0 := pose_trans(Wp0, p[0.02,0,0,0,0,0])
                        Wp := Wp0
                        Script: Wp[0]=ButtonPos[0]+0.01
                        Waypoint Variable (Variable): variable=Wp0
                        Waypoint Variable (Variable): variable=Wp
                        Set NoAction tcp=t4_Finger
                        Force Frame feature=Joint_6_name; selection=[0, 1, 1, 0, 0, 0]; wrench=[10, 20, -20, 0, 0, 0]; limitsForce=[0.01, 0.01, 0.025, 1.047198, 1.047198, 1.047198]; limitsMotion=[0.1, 0.1, 0.1, 0.349066, 0.349066, 0.349066]
                          Wait Sleep waitTime=1
                        Waypoint Variable (Variable): variable=Wp0
                      Folder Press down
                        Wp0 := pose_add(WpMultiringHi,Base_w_correctn)
                        Wp0 := pose_trans(Wp0, p[0.02,0,0,0,0,0])
                        Wp := Wp0
                        Script: Wp[0]=ButtonPos[0]+0.01
                        Waypoint Variable (Variable): variable=Wp0
                        Waypoint Variable (Variable): variable=Wp
                        Set NoAction tcp=t4_Finger
                        Force Frame feature=Joint_6_name; selection=[0, 1, 1, 0, 0, 0]; wrench=[10, 20, 20, 0, 0, 0]; limitsForce=[0.01, 0.01, 0.05, 1.047198, 1.047198, 1.047198]; limitsMotion=[0.1, 0.1, 0.1, 0.349066, 0.349066, 0.349066]
                          Wait Sleep waitTime=1
                        Waypoint Variable (Variable): variable=Wp0
                    Script: Report(2)
                  Else 
                    MoveJ speed 120 deg/s, acceleration 500 deg/s^2 (useActiveTCP=false positionType=JointAngles optimoveEnabled=false optiMoveSpeed=0.3 optiMoveAcceleration=0.09) tcp=t0_Flange; feature=Base
                      Waypoint WpBttnMidp: motionParameters(blendRadius=0.1); TCP in base x=-824.236 y=452.377 z=623.923 mm, rx=2.2214 ry=-2.2214 rz=0 rad; joints [161.838, -112.329, -68.535, -89.151, 90.318, 161.934] deg
                      Waypoint WpHome: TCP in base x=-539.74 y=192.879 z=621.496 mm, rx=3.1416 ry=0 rz=0 rad; joints [177.915, -76.399, -107.627, -86.021, 90.391, 88.106] deg
                    Script: Report(95)
            Folder 2W LMB FW
              If Progress_run()
                If In(ProgExe,[34])
                  SetCameraProg := 35
                  Timer (action=Reset) variable=T_Timeout
                  Timer (action=Start) variable=T_Timeout
                  Script: Report(13)
                  Wait Condition expression=Flags[3] or T_Timeout>60 or DEBUG or Abort
                  If Flags[3] or DEBUG
                    MoveL speed 1000 mm/s, acceleration 3000 mm/s^2 (useActiveTCP=false optimoveEnabled=false optiMoveSpeed=0.3 optiMoveAcceleration=0.09) tcp=t4_Finger; feature=Base
                      Folder Press FW
                        If False
                          Waypoint WpLmbFwMec: TCP in base x=-693.699 y=697.456 z=404.949 mm, rx=0.3536 ry=-3.0877 rz=0.0022 rad; joints [148.873, -132.515, -51.516, -84.507, 91.536, 225.911] deg; TCP offset x=-159 y=-58 z=70 mm, rx=0 ry=0 rz=0 rad
                        Wp := pose_add(WpLmbFwMec,Base_w_correctn)
                        Waypoint Variable (Variable): variable=Wp
                        Timer (action=Reset) variable=T_Timeout
                        Timer (action=Start) variable=T_Timeout
                        Force Frame feature=Joint_6_name; selection=[1, 0, 0, 0, 0, 0]; wrench=[-20, 10, -20, 0, 0, 0]; limitsForce=[0.05, 0.01, 0.05, 1.047198, 1.047198, 1.047198]; limitsMotion=[0.1, 0.1, 0.1, 0.349066, 0.349066, 0.349066]
                          Wait Condition expression=Flags[10] or T_Timeout>10 or (DEBUG and T_Timeout>2)
                        Waypoint Variable (Variable): variable=Wp
                  Else 
                    MoveJ speed 120 deg/s, acceleration 500 deg/s^2 (useActiveTCP=false positionType=JointAngles optimoveEnabled=false optiMoveSpeed=0.3 optiMoveAcceleration=0.09) tcp=t0_Flange; feature=Base
                      Waypoint WpBttnMidp: motionParameters(blendRadius=0.1); TCP in base x=-824.236 y=452.377 z=623.923 mm, rx=2.2214 ry=-2.2214 rz=0 rad; joints [161.838, -112.329, -68.535, -89.151, 90.318, 161.934] deg
                      Waypoint WpHome: TCP in base x=-539.74 y=192.879 z=621.496 mm, rx=3.1416 ry=0 rz=0 rad; joints [177.915, -76.399, -107.627, -86.021, 90.391, 88.106] deg
                    Script: Report(95)
            Folder 2W LMB RW
              If Progress_run()
                If In(ProgExe,[34])
                  Timer (action=Reset) variable=T_Timeout
                  Timer (action=Start) variable=T_Timeout
                  Script: Report(14)
                  Wait Condition expression=Flags[4] or T_Timeout>60 or DEBUG or Abort
                  If Flags[4] or DEBUG
                    MoveL speed 1000 mm/s, acceleration 3000 mm/s^2 (useActiveTCP=false optimoveEnabled=false optiMoveSpeed=0.3 optiMoveAcceleration=0.09) tcp=t4_Finger; feature=Base
                      Folder Press RW
                        If False
                          Waypoint WpLmbRwMec: TCP in base x=-698.526 y=711.31 z=401.685 mm, rx=0.3536 ry=-3.0877 rz=0.0022 rad; joints [148.396, -134.093, -49.101, -85.354, 91.549, 225.425] deg; TCP offset x=-159 y=-58 z=70 mm, rx=0 ry=0 rz=0 rad
                        Wp := pose_add(WpLmbRwMec,Base_w_correctn)
                        Waypoint Variable (Variable): variable=Wp
                        Timer (action=Reset) variable=T_Timeout
                        Timer (action=Start) variable=T_Timeout
                        Force Frame feature=Joint_6_name; selection=[1, 0, 0, 0, 0, 0]; wrench=[-20, 10, -20, 0, 0, 0]; limitsForce=[0.05, 0.01, 0.05, 1.047198, 1.047198, 1.047198]; limitsMotion=[0.1, 0.1, 0.1, 0.349066, 0.349066, 0.349066]
                          Wait Sleep waitTime=0.5
                        Force Frame feature=Joint_6_name; selection=[1, 0, 0, 0, 0, 0]; wrench=[-20, 10, -20, 0, 0, 0]; limitsForce=[0.01, 0.01, 0.05, 1.047198, 1.047198, 1.047198]; limitsMotion=[0.1, 0.1, 0.1, 0.349066, 0.349066, 0.349066]
                          Wait Condition expression=Flags[10] or T_Timeout>10 or (DEBUG and T_Timeout>2)
                        ButtonPos := get_actual_tcp_pose()
                        Waypoint Variable (Variable): variable=Wp
                  Else 
                    MoveJ speed 120 deg/s, acceleration 500 deg/s^2 (useActiveTCP=false positionType=JointAngles optimoveEnabled=false optiMoveSpeed=0.3 optiMoveAcceleration=0.09) tcp=t0_Flange; feature=Base
                      Waypoint WpBttnMidp: motionParameters(blendRadius=0.1); TCP in base x=-824.236 y=452.377 z=623.923 mm, rx=2.2214 ry=-2.2214 rz=0 rad; joints [161.838, -112.329, -68.535, -89.151, 90.318, 161.934] deg
                      Waypoint WpHome: TCP in base x=-539.74 y=192.879 z=621.496 mm, rx=3.1416 ry=0 rz=0 rad; joints [177.915, -76.399, -107.627, -86.021, 90.391, 88.106] deg
                    Script: Report(95)
            Folder Camera2
              If Progress_run()
                If In(ProgExe,[34])
                  SuppressedNode
                    SetCameraProg := 35
                  MoveL speed 1000 mm/s, acceleration 3000 mm/s^2 (useActiveTCP=false optimoveEnabled=false optiMoveSpeed=0.3 optiMoveAcceleration=0.09) tcp=t0_Flange; feature=Base
                    If False
                      Waypoint WpCamHeightUp: TCP in base x=-987.559 y=701.35 z=401.488 mm, rx=-0.4049 ry=3.1154 rz=0 rad; joints [152.865, -145.948, -34.796, -89.275, 90.298, 228.089] deg
                    Wp := pose_add(WpCamHeightUp,p[0,0,MeasHeight/1000,0,0,0])
                    SuppressedNode
                      Wp := WpCamHeightUp
                    Waypoint Variable (Variable): variable=Wp
                  Call CamAcquire
                  Script: CamData[1]=CamData[1]-MeasHeight/1000
                  Call CamCalculateCorectnPlane
            If Progress_run() and CamCorrectnOK≠ProgExe
              MoveJ speed 120 deg/s, acceleration 500 deg/s^2 (useActiveTCP=false optimoveEnabled=false optiMoveSpeed=0.3 optiMoveAcceleration=0.09) tcp=t0_Flange; feature=Base
                Waypoint WpBttnMidp: motionParameters(blendRadius=0.1); TCP in base x=-824.236 y=452.377 z=623.923 mm, rx=2.2214 ry=-2.2214 rz=0 rad; joints [161.838, -112.329, -68.535, -89.151, 90.318, 161.934] deg
                Waypoint WpHome: TCP in base x=-539.74 y=192.879 z=621.496 mm, rx=3.1416 ry=0 rz=0 rad; joints [177.915, -76.399, -107.627, -86.021, 90.391, 88.106] deg
              Script: Report(91)
            Folder Height up
              If Progress_run()
                If In(ProgExe,[34])
                  SetCameraProg := 36
                  Timer (action=Reset) variable=T_Timeout
                  Timer (action=Start) variable=T_Timeout
                  Script: Report(15)
                  Wait Condition expression=Flags[5] or T_Timeout>60 or DEBUG or Abort
                  If Flags[5] or DEBUG
                    MoveL speed 1000 mm/s, acceleration 3000 mm/s^2 (useActiveTCP=false optimoveEnabled=false optiMoveSpeed=0.3 optiMoveAcceleration=0.09) tcp=t4_Finger; feature=Base
                      Folder Press height up
                        If False
                          Waypoint WpHeiUp: TCP in base x=-696.215 y=774.447 z=367.033 mm, rx=0.2826 ry=-3.1275 rz=0.0033 rad; joints [145.509, -140.844, -40.709, -88.482, 90.438, 225.23] deg; TCP offset x=-159 y=-58 z=70 mm, rx=0 ry=0 rz=0 rad
                        Wp := pose_add(WpHeiUp,Base_w_correctn)
                        Script: Wp[0]=ButtonPos[0]-0.003
                        Waypoint Variable (Variable): variable=Wp
                        Set NoAction tcp=t4_Finger
                        Timer (action=Reset) variable=T_Timeout
                        Timer (action=Start) variable=T_Timeout
                        Force Frame feature=Base; selection=[0, 1, 1, 0, 0, 0]; wrench=[0, 0, 10, 0, 0, 0]; limitsForce=[0.02, 0.01, 0.05, 1.047198, 1.047198, 1.047198]; limitsMotion=[0.1, 0.1, 0.1, 0.349066, 0.349066, 0.349066]
                          Wait Condition expression=Flags[10] or T_Timeout>10 or (DEBUG and T_Timeout>2)
                        Wp0 := get_actual_tcp_pose()
                        Wp := pose_trans(Wp0, p[0.02,0,0.02,0,0,0])
                        Waypoint Variable (Variable): variable=Wp
                  Else 
                    MoveJ speed 120 deg/s, acceleration 500 deg/s^2 (useActiveTCP=false optimoveEnabled=false optiMoveSpeed=0.3 optiMoveAcceleration=0.09) tcp=t0_Flange; feature=Base
                      Waypoint WpBttnMidp: motionParameters(blendRadius=0.1); TCP in base x=-824.236 y=452.377 z=623.923 mm, rx=2.2214 ry=-2.2214 rz=0 rad; joints [161.838, -112.329, -68.535, -89.151, 90.318, 161.934] deg
                      Waypoint WpHome: TCP in base x=-539.74 y=192.879 z=621.496 mm, rx=3.1416 ry=0 rz=0 rad; joints [177.915, -76.399, -107.627, -86.021, 90.391, 88.106] deg
                    Script: Report(95)
            Folder Camera3
              If Progress_run()
                If In(ProgExe,[34])
                  SuppressedNode
                    SetCameraProg := 36
                  MoveL speed 1000 mm/s, acceleration 3000 mm/s^2 (useActiveTCP=false optimoveEnabled=false optiMoveSpeed=0.3 optiMoveAcceleration=0.09) tcp=t0_Flange; feature=Base
                    If False
                      Waypoint WpCamHeightDown: TCP in base x=-987.559 y=701.35 z=401.488 mm, rx=-0.4049 ry=3.1154 rz=0 rad; joints [152.865, -145.948, -34.796, -89.275, 90.298, 228.089] deg
                    Wp := pose_add(WpCamHeightUp,p[0,0,MeasHeight/1000,0,0,0])
                    SuppressedNode
                      Wp := WpCamHeightDown
                    Waypoint Variable (Variable): variable=Wp
                  Call CamAcquire
                  Script: CamData[1]=CamData[1]-MeasHeight/1000
                  Call CamCalculateCorectnPlane
            Folder Height down
              If Progress_run()
                If In(ProgExe,[34])
                  Timer (action=Reset) variable=T_Timeout
                  Timer (action=Start) variable=T_Timeout
                  Script: Report(16)
                  Wait Condition expression=Flags[6] or T_Timeout>60 or DEBUG or Abort
                  If Flags[6] or DEBUG
                    MoveL speed 1000 mm/s, acceleration 3000 mm/s^2 (useActiveTCP=false optimoveEnabled=false optiMoveSpeed=0.3 optiMoveAcceleration=0.09) tcp=t4_Finger; feature=Base
                      Folder Press height down
                        If False
                          Waypoint WpHeiDown: TCP in base x=-695.673 y=784.546 z=392.519 mm, rx=-0.3184 ry=3.1254 rz=0 rad; joints [145.284, -141.487, -36.989, -91.543, 90.3, 223.678] deg; TCP offset x=-159 y=-58 z=70 mm, rx=0 ry=0 rz=0 rad
                        Wp := pose_add(WpHeiDown,Base_w_correctn)
                        Script: Wp[0]=ButtonPos[0]-0.003
                        Wp0 := pose_add(Wp,p[-0.04,0,0,0,0,0])
                        Waypoint Variable (Variable): motionParameters(blendRadius=0.03); variable=Wp0
                        Waypoint Variable (Variable): variable=Wp
                        Set NoAction tcp=t4_Finger
                        Timer (action=Reset) variable=T_Timeout
                        Timer (action=Start) variable=T_Timeout
                        Force Frame feature=Base; selection=[0, 1, 1, 0, 0, 0]; wrench=[0, 0, -10, 0, 0, 0]; limitsForce=[0.02, 0.01, 0.05, 1.047198, 1.047198, 1.047198]; limitsMotion=[0.1, 0.1, 0.1, 0.349066, 0.349066, 0.349066]
                          Wait Condition expression=Flags[10] or T_Timeout>10
                        Wp := pose_trans(Wp, p[0.02,0,-0.02,0,0,0])
                        Waypoint Variable (Variable): variable=Wp
                    Script: Report(7)
                  Else 
                    MoveJ speed 120 deg/s, acceleration 500 deg/s^2 (useActiveTCP=false positionType=JointAngles optimoveEnabled=false optiMoveSpeed=0.3 optiMoveAcceleration=0.09) tcp=t0_Flange; feature=Base
                      Waypoint WpBttnMidp: motionParameters(blendRadius=0.1); TCP in base x=-824.236 y=452.377 z=623.923 mm, rx=2.2214 ry=-2.2214 rz=0 rad; joints [161.838, -112.329, -68.535, -89.151, 90.318, 161.934] deg
                      Waypoint WpHome: TCP in base x=-539.74 y=192.879 z=621.496 mm, rx=3.1416 ry=0 rz=0 rad; joints [177.915, -76.399, -107.627, -86.021, 90.391, 88.106] deg
                    Script: Report(95)
            If Progress_run()
              MoveJ speed 120 deg/s, acceleration 500 deg/s^2 (useActiveTCP=false positionType=JointAngles optimoveEnabled=false optiMoveSpeed=0.3 optiMoveAcceleration=0.09) tcp=t0_Flange; feature=Base
                Waypoint WpBttnMidp: motionParameters(blendRadius=0.1); TCP in base x=-824.236 y=452.377 z=623.923 mm, rx=2.2214 ry=-2.2214 rz=0 rad; joints [161.838, -112.329, -68.535, -89.151, 90.318, 161.934] deg
                Waypoint WpHome: TCP in base x=-539.74 y=192.879 z=621.496 mm, rx=3.1416 ry=0 rz=0 rad; joints [177.915, -76.399, -107.627, -86.021, 90.391, 88.106] deg
              Script: Report(50)
        Folder PushByHandle
          If In(ProgExe,[40])
            Script: Report(1)
            Folder AtHome? [hidden by the author, left out]
            SuppressedNode
              If Progress_run()
                SetCameraProg := 27
                MoveL speed 250 mm/s, acceleration 1200 mm/s^2 (useActiveTCP=false optimoveEnabled=false optiMoveSpeed=0.3 optiMoveAcceleration=0.09) tcp=t0_Flange; feature=Base
                  Waypoint WpBttnMidp1: motionParameters(blendRadius=0.1); TCP in base x=-465.361 y=283.426 z=636.73 mm, rx=-2.2214 ry=2.2214 rz=0 rad; joints [167.185, -73.405, -108.257, -88.385, 90.398, 167.36] deg
                  Waypoint WpBttnMidp2: motionParameters(blendRadius=0.1); TCP in base x=-296.641 y=583.561 z=625.265 mm, rx=-1.2596 ry=2.878 rz=0 rad; joints [132.275, -84.542, -100.549, -84.955, 90.381, 175.201] deg
                  Waypoint WpBttnMidp3: motionParameters(blendRadius=0.1); TCP in base x=114.747 y=708.142 z=644.758 mm, rx=0 ry=3.1416 rz=0 rad; joints [94.755, -90.505, -92.903, -86.639, 90.379, 184.947] deg; TCP offset x=0 y=0 z=0 mm, rx=0 ry=0 rz=0 rad
                  Waypoint WpCamLMB: TCP in base x=186.376 y=644.645 z=421.712 mm, rx=0.3238 ry=3.0539 rz=-0.0115 rad; joints [89.517, -91.476, -115.043, -64.369, 86.327, 191.973] deg
                Call CamAcquire
                CamCorrection := p[0,CamData[0],CamData[1],0,0,0]
            SuppressedNode
              If Progress_run() and CamCorrectnOK≠ProgExe
                MoveL speed 250 mm/s, acceleration 1200 mm/s^2 (useActiveTCP=false optimoveEnabled=false optiMoveSpeed=0.3 optiMoveAcceleration=0.09) tcp=t0_Flange; feature=Base
                  Waypoint WpBttnMidp3: motionParameters(blendRadius=0.1); TCP in base x=114.747 y=708.142 z=644.758 mm, rx=0 ry=3.1416 rz=0 rad; joints [94.755, -90.505, -92.903, -86.639, 90.379, 184.947] deg; TCP offset x=0 y=0 z=0 mm, rx=0 ry=0 rz=0 rad
                  Waypoint WpBttnMidp2: motionParameters(blendRadius=0.1); TCP in base x=-296.641 y=583.561 z=625.265 mm, rx=-1.2596 ry=2.878 rz=0 rad; joints [132.275, -84.542, -100.549, -84.955, 90.381, 175.201] deg
                  Waypoint WpBttnMidp1: motionParameters(blendRadius=0.1); TCP in base x=-465.361 y=283.426 z=636.73 mm, rx=-2.2214 ry=2.2214 rz=0 rad; joints [167.185, -73.405, -108.257, -88.385, 90.398, 167.36] deg
                  Waypoint WpHome: TCP in base x=-539.74 y=192.879 z=621.496 mm, rx=3.1416 ry=0 rz=0 rad; joints [177.915, -76.399, -107.627, -86.021, 90.391, 88.106] deg
                Script: Report(91)
            If Progress_run() and  not AdapterDocked
              Script: Report(94)
            If Progress_run()
              PusherReturn := False
              Set DigitalOutput pin=Do_PusherReturn; digitalValue=0
              Set DigitalOutput pin=Do_PusherWork; digitalValue=1
              Wait Condition expression=PusherPosStable and PusherPosDev>-20
              Set DigitalOutput pin=Do_PusherWork; digitalValue=0
              Call GripperOpen
              Set NoAction tcp=t2_Gripper
              MoveL speed 1000 mm/s, acceleration 3000 mm/s^2 (useActiveTCP=false optimoveEnabled=false optiMoveSpeed=0.3 optiMoveAcceleration=0.09) tcp=t2_Gripper; feature=Base
                Waypoint WpHandle0: motionParameters(blendRadius=0.05); TCP in base x=-444.611 y=570.363 z=233.755 mm, rx=3.1416 ry=0 rz=0 rad; joints [163.57, -85.97, -134.254, -49.795, 90.223, 73.938] deg; TCP offset x=0 y=-260 z=74 mm, rx=0 ry=0 rz=0 rad
                Waypoint WpHandle: TCP in base x=-407.419 y=672.326 z=245.413 mm, rx=3.1416 ry=0 rz=0 rad; joints [151.912, -88.862, -130.027, -51.129, 90.225, 62.271] deg
                Force Frame feature=Joint_6_name; selection=[0, 1, 0, 0, 0, 0]; wrench=[0, -10, 0, 0, 0, 0]; limitsForce=[0.15, 0.05, 0.15, 1.047198, 1.047198, 1.047198]; limitsMotion=[0.1, 0.1, 0.1, 0.349066, 0.349066, 0.349066]
                  Wait Sleep waitTime=1
                Force Frame feature=Joint_6_name; selection=[0, 1, 1, 0, 0, 0]; wrench=[0, -10, -80, 0, 0, 0]; limitsForce=[0.15, 0.05, 0.05, 1.047198, 1.047198, 1.047198]; limitsMotion=[0.1, 0.1, 0.1, 0.349066, 0.349066, 0.349066]
                  Wait Sleep waitTime=1
                Force Frame feature=Joint_6_name; selection=[0, 1, 1, 0, 0, 0]; wrench=[0, -30, -80, 0, 0, 0]; limitsForce=[0.15, 0.5, 0.05, 1.047198, 1.047198, 1.047198]; limitsMotion=[0.1, 0.1, 0.1, 0.349066, 0.349066, 0.349066]
                  Wait Sleep waitTime=0.2
                  Set DigitalOutput pin=Do_PusherReturn; digitalValue=0
                  Set DigitalOutput pin=Do_PusherWork; digitalValue=1
                  Wait AnalogInput pin=analog_in[0]; analogComparison=0; analogValue=8.5
                  Wait Sleep waitTime=2
                  Set DigitalOutput pin=Do_PusherWork; digitalValue=0
                PusherReturn := True
                Waypoint WpOffHandle (Relative): relativeFromPosition TCP in base x=-402.966 y=514.879 z=380.999 mm, rx=3.1271 ry=-0.0003 rz=-0.0016 rad; joints [143.175, -92.106, -119.096, -59.265, 90.96, 53.495] deg; TCP in base x=-408.771 y=503.734 z=306.943 mm, rx=3.132 ry=-0.0002 rz=0.0026 rad; joints [144.358, -96.318, -123.61, -50.484, 90.601, 54.716] deg
                Waypoint WpHandle0: TCP in base x=-444.611 y=570.363 z=233.755 mm, rx=3.1416 ry=0 rz=0 rad; joints [163.57, -85.97, -134.254, -49.795, 90.223, 73.938] deg; TCP offset x=0 y=-260 z=74 mm, rx=0 ry=0 rz=0 rad
              MoveL speed 1000 mm/s, acceleration 3000 mm/s^2 (useActiveTCP=false optimoveEnabled=false optiMoveSpeed=0.3 optiMoveAcceleration=0.09) tcp=t0_Flange; feature=Base
                Waypoint WpHome: TCP in base x=-539.74 y=192.879 z=621.496 mm, rx=3.1416 ry=0 rz=0 rad; joints [177.915, -76.399, -107.627, -86.021, 90.391, 88.106] deg
              Script: Report(50)
        Folder Tilt manual adjust
          If In(ProgExe,[42])
            Script: Report(1)
            Folder AtHome? [hidden by the author, left out]
            If Progress_run() and  not AdapterDocked
              Script: Report(94)
            If Progress_run()
              Set NoAction tcp=t2_Gripper
              ''
              If InRange(Tilt_PV-CMD_Tilt_SP,-60,60)
                'Laser value in range'
                MaxTiltPumps := 10
                If InRange(Tilt_PV-CMD_Tilt_SP,-60,-3)
                  'Tilt too high'
                  Call GripperClose
                  MoveJ speed 120 deg/s, acceleration 500 deg/s^2 (useActiveTCP=false positionType=JointAngles optimoveEnabled=false optiMoveSpeed=0.3 optiMoveAcceleration=0.09) tcp=t2_Gripper; feature=Base
                    Waypoint WpTilt0: motionParameters(blendRadius=0.05); TCP in base x=-227.69 y=551.131 z=582.792 mm, rx=2.0545 ry=-0.3038 rz=1.9788 rad; joints [159.442, -91.98, -95.337, -171.039, 89.315, 86.776] deg; TCP offset x=0 y=-260 z=74 mm, rx=0 ry=0 rz=0 rad
                    Waypoint WpTilt1: motionParameters(blendRadius=0.05); TCP in base x=-257.589 y=472.823 z=277.035 mm, rx=1.2192 ry=1.1986 rz=1.2029 rad; joints [148.759, -96.668, -96.779, -166.311, 59.701, -0.146] deg
                    Waypoint WpTiltDown: TCP in base x=-255.62 y=660.561 z=224.593 mm, rx=1.6089 ry=0.8926 rz=1.5881 rad; joints [144.727, -102.698, -98.998, -157.618, 55.587, 30.735] deg; TCP offset x=0 y=-260 z=74 mm, rx=0 ry=0 rz=0 rad
                    Force Frame feature=Joint_6_name; selection=[1, 1, 0, 0, 0, 0]; wrench=[15, 0, 0, 0, 0, 0]; limitsForce=[0.1, 0.15, 0.15, 1.047198, 1.047198, 1.047198]; limitsMotion=[0.1, 0.1, 0.1, 0.349066, 0.349066, 0.349066]
                      Wait Sleep waitTime=1
                    Wp := P_act
                    Loop While (checkContinuously=false) expression=InRange(Tilt_PV-CMD_Tilt_SP,-60,-5) and MaxTiltPumps>0
                      Force Frame feature=Joint_6_name; selection=[1, 1, 0, 0, 0, 0]; wrench=[10, -100, 0, 0, 0, 0]; limitsForce=[0.15, 0.1, 0.15, 1.047198, 1.047198, 1.047198]; limitsMotion=[0.1, 0.1, 0.1, 0.349066, 0.349066, 0.349066]
                        Wait Sleep waitTime=1.5
                      Waypoint Variable (Variable): variable=Wp
                      MaxTiltPumps := MaxTiltPumps-1
                    Waypoint WpTiltDown: motionParameters(blendRadius=0.05); TCP in base x=-255.62 y=660.561 z=224.593 mm, rx=1.6089 ry=0.8926 rz=1.5881 rad; joints [144.727, -102.698, -98.998, -157.618, 55.587, 30.735] deg
                    Waypoint WpTilt1: motionParameters(blendRadius=0.05); TCP in base x=-257.589 y=472.823 z=277.035 mm, rx=1.2192 ry=1.1986 rz=1.2029 rad; joints [148.759, -96.668, -96.779, -166.311, 59.701, -0.146] deg; TCP offset x=0 y=-260 z=74 mm, rx=0 ry=0 rz=0 rad
                    Waypoint WpTilt0: TCP in base x=-227.69 y=551.131 z=582.792 mm, rx=2.0545 ry=-0.3038 rz=1.9788 rad; joints [159.442, -91.98, -95.337, -171.039, 89.315, 86.776] deg
                  MoveJ speed 120 deg/s, acceleration 500 deg/s^2 (useActiveTCP=false positionType=JointAngles optimoveEnabled=false optiMoveSpeed=0.3 optiMoveAcceleration=0.09) tcp=t0_Flange; feature=Base
                    Waypoint WpHome: TCP in base x=-539.74 y=192.879 z=621.496 mm, rx=3.1416 ry=0 rz=0 rad; joints [177.915, -76.399, -107.627, -86.021, 90.391, 88.106] deg
                ElseIf InRange(Tilt_PV-CMD_Tilt_SP,3,60)
                  'Tilt too low'
                  Call GripperClose
                  MoveJ speed 120 deg/s, acceleration 500 deg/s^2 (useActiveTCP=false positionType=JointAngles optimoveEnabled=false optiMoveSpeed=0.3 optiMoveAcceleration=0.09) tcp=t2_Gripper; feature=Base
                    Waypoint WpTilt0: motionParameters(blendRadius=0.05); TCP in base x=-227.69 y=551.131 z=582.792 mm, rx=2.0545 ry=-0.3038 rz=1.9788 rad; joints [159.442, -91.98, -95.337, -171.039, 89.315, 86.776] deg; TCP offset x=0 y=-260 z=74 mm, rx=0 ry=0 rz=0 rad
                    Waypoint WpTilt1: motionParameters(blendRadius=0.05); TCP in base x=-257.589 y=472.823 z=277.035 mm, rx=1.2192 ry=1.1986 rz=1.2029 rad; joints [148.759, -96.668, -96.779, -166.311, 59.701, -0.146] deg
                    Waypoint WpTiltUp: TCP in base x=-252.613 y=628.413 z=253.114 mm, rx=1.2758 ry=1.1614 rz=1.2589 rad; joints [139.268, -106.731, -87.005, -165.884, 50.193, 4.176] deg; TCP offset x=0 y=-260 z=74 mm, rx=0 ry=0 rz=0 rad
                    Force Frame feature=Joint_6_name; selection=[1, 1, 0, 0, 0, 0]; wrench=[15, 0, 0, 0, 0, 0]; limitsForce=[0.1, 0.15, 0.15, 1.047198, 1.047198, 1.047198]; limitsMotion=[0.1, 0.1, 0.1, 0.349066, 0.349066, 0.349066]
                      Wait Sleep waitTime=1
                    Wp := P_act
                    Loop While (checkContinuously=false) expression=InRange(Tilt_PV-CMD_Tilt_SP,5,60) and MaxTiltPumps>0
                      Force Frame feature=Joint_6_name; selection=[1, 1, 0, 0, 0, 0]; wrench=[10, 100, 0, 0, 0, 0]; limitsForce=[0.15, 0.1, 0.15, 1.047198, 1.047198, 1.047198]; limitsMotion=[0.1, 0.1, 0.1, 0.349066, 0.349066, 0.349066]
                        Wait Sleep waitTime=1.5
                      Waypoint Variable (Variable): variable=Wp
                      MaxTiltPumps := MaxTiltPumps-1
                    Waypoint WpTiltUp: motionParameters(blendRadius=0.05); TCP in base x=-252.613 y=628.413 z=253.114 mm, rx=1.2758 ry=1.1614 rz=1.2589 rad; joints [139.268, -106.731, -87.005, -165.884, 50.193, 4.176] deg
                    Waypoint WpTilt1: motionParameters(blendRadius=0.05); TCP in base x=-257.589 y=472.823 z=277.035 mm, rx=1.2192 ry=1.1986 rz=1.2029 rad; joints [148.759, -96.668, -96.779, -166.311, 59.701, -0.146] deg; TCP offset x=0 y=-260 z=74 mm, rx=0 ry=0 rz=0 rad
                    Waypoint WpTilt0: motionParameters(blendRadius=0.05); TCP in base x=-227.69 y=551.131 z=582.792 mm, rx=2.0545 ry=-0.3038 rz=1.9788 rad; joints [159.442, -91.98, -95.337, -171.039, 89.315, 86.776] deg
                    Waypoint WpHome: TCP in base x=-539.74 y=192.879 z=621.496 mm, rx=3.1416 ry=0 rz=0 rad; joints [177.915, -76.399, -107.627, -86.021, 90.391, 88.106] deg
              Else 
                Script: Report(93)
              Script: Report(50)
        Folder Program finished
          ProgDn := ProgExe
          ProgExe := 0
      Folder Parking
        If Parking≟10 or ProgExe≟1011
          Wait Condition expression=EvtDock≤0
          If AtHomePos
            MoveJ speed 120 deg/s, acceleration 500 deg/s^2 (useActiveTCP=true positionType=JointAngles optimoveEnabled=false optiMoveSpeed=0.3 optiMoveAcceleration=0.09) feature=Base
              Waypoint WpPark: TCP in base x=-21.021 y=216.43 z=1228.484 mm, rx=-2.2794 ry=-2.1557 rz=0.0038 rad; joints [148.842, -80.043, -21.696, -168.004, 90.169, -28.26] deg
              STS_Reservation := 0
          Parking := 0
          If DEBUG
            ProgExe := 0
        If Parking≟1 or ProgExe≟1001
          If AtParkPos
            MoveJ speed 120 deg/s, acceleration 500 deg/s^2 (useActiveTCP=true positionType=JointAngles optimoveEnabled=false optiMoveSpeed=0.3 optiMoveAcceleration=0.09) feature=Base
              Waypoint WpHome: TCP in base x=-539.74 y=192.879 z=621.496 mm, rx=3.1416 ry=0 rz=0 rad; joints [177.915, -76.399, -107.627, -86.021, 90.391, 88.106] deg
              STS_Reservation := 1
            Parking := 0
            If DEBUG
              ProgExe := 0
  Script: sync()
Thread Thread_1 (runOnlyOnce=false)
  Folder Continuous calculations
    Folder get live force and tcp pos
      P_act := get_actual_tcp_pose()
      V_act := get_actual_tcp_speed()
      V_act_norm := norm(V_act)
      ToolForce := norm(get_tcp_force())
      P_Flange := get_actual_tool_flange_pose()
      D_rel := pose_sub(P_act, P_ini)
      AtHomePos := pose_dist(P_Flange, WpHome)<0.005
      AtParkPos := pose_dist(P_Flange, WpPark)<0.005
      AdapterDocked := Di_Docked
      Tilt_PV := (Ai_LaserTilt*100+505)*0.1+Tilt_PV*0.9
      Folder Calculate actual offset in tool frame
        If ProgExe≟15
          TempWp := pose_sub(WpBuckleSpa1,Base_w_correctn)
          BklToolDist := pose_trans(pose_inv(TempWp), P_act)
        If ProgExe≟16
          TempWp := pose_sub(WpBuckleSpa3,Base_w_correctn)
          BklToolDist := pose_trans(pose_inv(TempWp), P_act)
      Folder InterlockOutput
        If P_Flange[1]>-0.45
          Set DigitalOutput pin=Do_SafePosition; digitalValue=1
        ElseIf P_Flange[0]>0
          Set DigitalOutput pin=Do_SafePosition; digitalValue=1
        Else 
          Set DigitalOutput pin=Do_SafePosition; digitalValue=0
    Folder Modbus mapping
      Folder Heartbeat
        Timer (action=Start) variable(name=T_Heartbeat)
        If T_Heartbeat≥1
          Timer (action=Reset) variable=T_Heartbeat
          If STS_Heartbeat
            STS_Heartbeat := False
          Else 
            STS_Heartbeat := True
      Folder Safe position
        STS_Safe := True
        If pose_dist(P_act,WpBuckleSpa1)<0.2
          STS_Safe := False
        If pose_dist(P_act,WpConnSpa1EL)<0.08
          STS_Safe := False
        If pose_dist(P_act,WpHandle)<0.08
          STS_Safe := False
        If pose_dist(P_act,WpHeiUp)<0.08
          STS_Safe := False
        If pose_dist(P_act,WpLmbFwEL)<0.08
          STS_Safe := False
        If pose_dist(P_act,WpUnplug1_3)<0.08
          STS_Safe := False
        If pose_dist(P_act,WpUnplg1_3M)<0.08
          STS_Safe := False
      Folder Outputs
        Script: write_port_register(129,STS_Progress)
        Script: write_port_register(131,STS_Reservation)
        Script: write_port_register(134,binary_list_to_integer ([digital_in[0], False ,config_in[0],STS_Heartbeat,STS_Safe, False ]))
      Folder Inputs
        CMD_Reserve_i1 := read_port_register(160)
        CMD_Timeout_i1 := read_port_register(162)
        CMD_Program_i1 := read_port_register(164)
        CMD_Tilt_SP := read_port_register(166)
        CMD_Flags_i1 := read_port_register(170)
        CMD_Heartbt_i1 := read_port_register(180)
      Folder Generate flags
        Flags := integer_to_binary_list(CMD_Flags_i1)
    Folder Speed
      Timer (action=Start) variable(name=T_SpeedSet)
      If T_SpeedSet>2 and  not DEBUG
        Script: socket_send_string("set speed")
        Script: socket_send_string(1)
        Script: socket_send_byte(10)
        Timer (action=Reset) variable=T_SpeedSet
    Wait Sleep waitTime=0.01
  Folder ReservationControl
    If STS_Reservation≟0 and ProgExe≟0
      If CMD_Reserve_i1≟1
        'request reservation'
        If AtHomePos or AdapterReady
          STS_Reservation := 1
        Else 
          Parking := 1
    'Timeout reservation - station keeps reservation for a while to prevent other app stealing the process'
    'Timeout is configurable, so application can control how long to keep robot before letting other app'
    If STS_Progress≟0 and STS_Reservation≠0
      If STS_Reservation≟1 and CMD_Reserve_i1≟1
        'nop'
      Else 
        T_KeepReservtn := CMD_Timeout_i1
        Timer (action=Start) variable(name=tim_Unreserve)
        If tim_Unreserve>T_KeepReservtn
          STS_Reservation := 0
          Timer (action=Stop) variable=tim_Unreserve
    Else 
      Timer (action=Stop) variable=tim_Unreserve
      Timer (action=Reset) variable=tim_Unreserve
    'Force release reservation from app - in case of intervetion'
    If STS_Progress≟0 and In(STS_Reservation,[0,1]) and In(CMD_Reserve_i1,[98,99]) and  not DEBUG
      If AtHomePos
        Parking := 10
      If AtParkPos
        STS_Reservation := 0
      If CMD_Reserve_i1≟99 and  not Mute
        Set DigitalOutput pin=Do_Blue; digitalValue=1
        Set DigitalOutput pin=Do_Horn; digitalValue=1
    Wait Sleep waitTime=0.01
  Folder Program control
    'Start new Prog / Confirm Prog Running'
    If STS_Progress≟0 and ProgExe≟0  and  not Abort and  not DEBUG
      If InRange(CMD_Program_i1,10,49) and STS_Reservation≟1
        ProgExe := CMD_Program_i1
        T_KeepReservtn := CMD_Timeout_i1
        Script: Report(0)
    'Ack results - get ready for new prg'
    If ProgExe≟0 and Progress_finished()
      If CMD_Program_i1≠ProgDn
        STS_Progress := 0
  Folder Pusher Control
    If PusherReturn and NormalMode
      Set DigitalOutput pin=Do_PusherReturn; digitalValue=1
      Set DigitalOutput pin=Do_PusherWork; digitalValue=0
      Timer (action=Start) variable(name=T_Pusher)
      If T_Pusher>20 or Di_Pusher_Bp
        Set DigitalOutput pin=Do_PusherReturn; digitalValue=0
        PusherReturn := False
    Else 
      Timer (action=Stop) variable=T_Pusher
      Timer (action=Reset) variable=T_Pusher
    If not NormalMode
      Set DigitalOutput pin=Do_PusherReturn; digitalValue=0
      Set DigitalOutput pin=Do_PusherWork; digitalValue=0
    If Flags[11] and NormalMode
      'Activate pusher in advance'
      Set DigitalOutput pin=Do_PusherReturn; digitalValue=0
      Set DigitalOutput pin=Do_PusherWork; digitalValue=1
    PusherPos := Calibrate(Ai_Pusher,1,8,260,385)
    PusherPosFt := PusherPos*0.2+PusherPosFt*0.8
    PusherPosStable := InRange(PusherPosFt-PusherPos,-1,1) and PusherPosFt>265
  Folder Operator call deactivation
    If Do_Blue or Do_Horn
      Timer (action=Start) variable(name=T_Call)
      If not  NormalMode and T_Call>4
        Set DigitalOutput pin=Do_Blue; digitalValue=0
        Set DigitalOutput pin=Do_Horn; digitalValue=0
        Mute := True
    Else 
      Timer (action=Stop) variable=T_Call
      Timer (action=Reset) variable=T_Call
  Folder Abort
    If Flags[14]
      Abort := True
    If AtHomePos or AtParkPos
      Abort := False
    If Abort
      If AdapterReady
        EvtDock := 1
  Wait Sleep waitTime=0.01
SubProgram WaitForNormalMode [hidden by the author, left out]
SubProgram  [hidden by the author, left out]
SubProgram  [hidden by the author, left out]
SubProgram  [hidden by the author, left out]
SubProgram  [hidden by the author, left out]
Event  expression=SetCameraProg>0
  Folder Set program to camera in advance
    Set DigitalOutput pin=CnxDO_Trig; digitalValue=0
    Set DigitalOutput pin=CnxDO_TrigEn; digitalValue=1
    Script: modbus_delete_signal("CnxAO_Program")
    Script: modbus_add_signal("192.168.1.101", 255, 2001, 16, "CnxAO_Program", True ,1)
    Script: modbus_set_output_register("CnxAO_Program",SetCameraProg, False )
    Wait Sleep waitTime=0.2
    Set DigitalOutput pin=CnxDO_SetUsrDta; digitalValue=1
    Wait DigitalInput pin=CnxDi_UsrDtaAck; digitalValue=1
    Set DigitalOutput pin=CnxDO_SetUsrDta; digitalValue=0
    Set DigitalOutput pin=CnxDO_SoftEvt0; digitalValue=1
    Wait DigitalInput pin=CnxDI_Evt0Ack; digitalValue=1
    Set DigitalOutput pin=CnxDO_SoftEvt0; digitalValue=0
    Timer (action=Reset) variable=CamTimeout
    Timer (action=Start) variable=CamTimeout
    Wait Condition expression=CnxAI_Program≟SetCameraProg or CamTimeout>3
    If CnxAI_Program≠SetCameraProg
      Folder For the first time it needs trigger when going online
        Set DigitalOutput pin=CnxDO_Trig; digitalValue=1
        Wait Sleep waitTime=1
        Set DigitalOutput pin=CnxDO_Trig; digitalValue=0
        Script: textmsg("extra cam trigger on program set")
      If CnxAI_Program≠SetCameraProg
        SuppressedNode
          Popup Error (haltProgram=false message=Error: camera program not set inputType=Text)
      Else 
        Wait Sleep waitTime=0.5
        SetCameraProg := 0
    Else 
      Wait Sleep waitTime=0.5
      SetCameraProg := 0
  If SetCameraProg>0
    'repeat on fail'
    Wait Sleep waitTime=3
    Folder Set program to camera in advance
      Set DigitalOutput pin=CnxDO_Trig; digitalValue=0
      Set DigitalOutput pin=CnxDO_TrigEn; digitalValue=1
      Script: modbus_delete_signal("CnxAO_Program")
      Script: modbus_add_signal("192.168.1.101", 255, 2001, 16, "CnxAO_Program", True ,1)
      Script: modbus_set_output_register("CnxAO_Program",SetCameraProg, False )
      Wait Sleep waitTime=0.2
      Set DigitalOutput pin=CnxDO_SetUsrDta; digitalValue=1
      Wait DigitalInput pin=CnxDi_UsrDtaAck; digitalValue=1
      Set DigitalOutput pin=CnxDO_SetUsrDta; digitalValue=0
      Set DigitalOutput pin=CnxDO_SoftEvt0; digitalValue=1
      Wait DigitalInput pin=CnxDI_Evt0Ack; digitalValue=1
      Set DigitalOutput pin=CnxDO_SoftEvt0; digitalValue=0
      Timer (action=Reset) variable=CamTimeout
      Timer (action=Start) variable=CamTimeout
      Wait Condition expression=CnxAI_Program≟SetCameraProg or CamTimeout>3
      If CnxAI_Program≠SetCameraProg
        Folder For the first time it needs trigger when going online
          Set DigitalOutput pin=CnxDO_Trig; digitalValue=1
          Wait Sleep waitTime=1
          Set DigitalOutput pin=CnxDO_Trig; digitalValue=0
          Script: textmsg("extra cam trigger on program set")
        If CnxAI_Program≠SetCameraProg
          SuppressedNode
            Popup Error (haltProgram=false message=Error: camera program not set inputType=Text)
        Else 
          Wait Sleep waitTime=0.5
          SetCameraProg := 0
      Else 
        Wait Sleep waitTime=0.5
        SetCameraProg := 0
  If SetCameraProg>0
    'repeat on fail'
    Wait Sleep waitTime=3
    Folder Set program to camera in advance
      Set DigitalOutput pin=CnxDO_Trig; digitalValue=0
      Set DigitalOutput pin=CnxDO_TrigEn; digitalValue=1
      Script: modbus_delete_signal("CnxAO_Program")
      Script: modbus_add_signal("192.168.1.101", 255, 2001, 16, "CnxAO_Program", True ,1)
      Script: modbus_set_output_register("CnxAO_Program",SetCameraProg, False )
      Wait Sleep waitTime=0.2
      Set DigitalOutput pin=CnxDO_SetUsrDta; digitalValue=1
      Wait DigitalInput pin=CnxDi_UsrDtaAck; digitalValue=1
      Set DigitalOutput pin=CnxDO_SetUsrDta; digitalValue=0
      Set DigitalOutput pin=CnxDO_SoftEvt0; digitalValue=1
      Wait DigitalInput pin=CnxDI_Evt0Ack; digitalValue=1
      Set DigitalOutput pin=CnxDO_SoftEvt0; digitalValue=0
      Timer (action=Reset) variable=CamTimeout
      Timer (action=Start) variable=CamTimeout
      Wait Condition expression=CnxAI_Program≟SetCameraProg or CamTimeout>3
      If CnxAI_Program≠SetCameraProg
        Folder For the first time it needs trigger when going online
          Set DigitalOutput pin=CnxDO_Trig; digitalValue=1
          Wait Sleep waitTime=1
          Set DigitalOutput pin=CnxDO_Trig; digitalValue=0
          Script: textmsg("extra cam trigger on program set")
        If CnxAI_Program≠SetCameraProg
          SuppressedNode
            Popup Error (haltProgram=false message=Error: camera program not set inputType=Text)
        Else 
          Wait Sleep waitTime=0.5
          SetCameraProg := 0
      Else 
        Wait Sleep waitTime=0.5
        SetCameraProg := 0
  If SetCameraProg>0
    Popup Error (haltProgram=false message=Error: camera program not set inputType=Text)
SubProgram -> CamAcquire
SubProgram -> CamCalculateCorectnPlane
Event  expression=EvtDock>0
  Folder Dock
    MoveL speed 1000 mm/s, acceleration 3000 mm/s^2 (useActiveTCP=false optimoveEnabled=false optiMoveSpeed=0.3 optiMoveAcceleration=0.09) tcp=t2_Gripper; feature=Base
      If EvtDock≟2
        Folder Force mvts
          Set NoAction tcp=t2_Gripper
          Wp0 := P_act
          Force Frame feature=Joint_6_name; selection=[0, 1, 0, 0, 0, 0]; wrench=[0, -20, 0, 0, 0, 0]; limitsForce=[0.15, 0.1, 0.15, 1.047198, 1.047198, 1.047198]; limitsMotion=[0.1, 0.1, 0.1, 0.349066, 0.349066, 0.349066]
            Wait Sleep waitTime=1
          Force Frame feature=Joint_6_name; selection=[1, 0, 1, 0, 0, 0]; wrench=[0, -10, 0, 0, 0, 0]; limitsForce=[0.15, 0.05, 0.1, 1.047198, 1.047198, 1.047198]; limitsMotion=[0.1, 0.1, 0.1, 0.349066, 0.349066, 0.349066]
            Wait Sleep waitTime=0.2
            Call GripperClose
            Wait Sleep waitTime=0.2
          If timer_Gripper>3
            Call GripperOpen
            MoveL speed 500 mm/s, acceleration 1200 mm/s^2 (useActiveTCP=true optimoveEnabled=false optiMoveSpeed=0.3 optiMoveAcceleration=0.09) feature=Base
              Waypoint Variable (Variable): variable=Wp0
            Force Frame feature=Joint_6_name; selection=[0, 1, 0, 0, 0, 0]; wrench=[0, -20, 0, 0, 0, 0]; limitsForce=[0.15, 0.1, 0.15, 1.047198, 1.047198, 1.047198]; limitsMotion=[0.1, 0.1, 0.1, 0.349066, 0.349066, 0.349066]
              Wait Sleep waitTime=1
            Force Frame feature=Joint_6_name; selection=[1, 0, 1, 0, 0, 0]; wrench=[0, -10, 0, 0, 0, 0]; limitsForce=[0.15, 0.05, 0.1, 1.047198, 1.047198, 1.047198]; limitsMotion=[0.1, 0.1, 0.1, 0.349066, 0.349066, 0.349066]
              Wait Sleep waitTime=0.2
              Call GripperClose
              Wait Sleep waitTime=0.2
          If timer_Gripper>3
            Call GripperOpen
            MoveL speed 500 mm/s, acceleration 1200 mm/s^2 (useActiveTCP=true optimoveEnabled=false optiMoveSpeed=0.3 optiMoveAcceleration=0.09) feature=Base
              Waypoint Variable (Variable): variable=Wp0
              EvtDock := -97
          If EvtDock≟2
            MoveDirectionNode (selectedDirection=YPlus) feature=Joint_6_name
              Until DISTANCE (allowActions=false deceleration=3 distanceNodeType=BLEND) Distance=0.1; motionParameters(blendRadius=0.04)
      If EvtDock>0
        Script: Report(40)
        Wp := pose_trans(WpDock, p[0,0.25,0,0,0,0])
        Waypoint Variable (Variable): motionParameters(blendRadius=0.05); variable=Wp
        Waypoint WpDock referenceName=WpDock: TCP in base x=-85.659 y=314.493 z=77.7 mm, rx=1.8875 ry=-1.8567 rz=-0.5938 rad; joints [149.519, -78.77, -155.163, -4.834, 107.001, 153.83] deg
        Call GripperOpen
        Waypoint Variable (Variable): variable=Wp
        MoveL speed 1000 mm/s, acceleration 3000 mm/s^2 (useActiveTCP=false optimoveEnabled=false optiMoveSpeed=0.3 optiMoveAcceleration=0.09) tcp=t0_Flange; feature=Base
          Waypoint WpHome: TCP in base x=-539.74 y=192.879 z=621.496 mm, rx=3.1416 ry=0 rz=0 rad; joints [177.915, -76.399, -107.627, -86.021, 90.391, 88.106] deg
        EvtDock := 0
    AdapterReady := False
Event  expression=EvtBeep
  Loop While (checkContinuously=false) expression=EvtBeep
    Set DigitalOutput pin=Do_Horn; digitalValue=1
    Set DigitalOutput pin=Do_Blue; digitalValue=1
    Wait Sleep waitTime=0.5
    Set DigitalOutput pin=Do_Horn; digitalValue=0
    Set DigitalOutput pin=Do_Blue; digitalValue=0
    Wait Sleep waitTime=5
SubProgram GripperOpen [hidden by the author, left out]
SubProgram GripperOpenQuick [hidden by the author, left out]
SubProgram GripperClose [hidden by the author, left out]
SubProgram CamAcquire (keepSynchronizedWithDisk=false)
  Folder Trig camera and process data [hidden by the author, left out]
SubProgram GripperCloseQuick [hidden by the author, left out]
SubProgram CamCalculateCorectnPlane (keepSynchronizedWithDisk=false)
  Folder Folder [hidden by the author, left out]
